(* IEC 61131-3 sources: Lasal-MCP/examples/SampleSource/LASALScreenAdvancedSolution/LASALScreenAdvancedSolution/LASALScreenAdvacnedSolution/Stations/Terminal/HMI/Class/InputMyIO, 1 file *)

(* ---- InputMyIO.st ---- *)
#define CROSSHAIR_LENGTH 20
#define CROSSHAIR_WIDTH 1
#define OFFSET_X 10
#define OFFSET_Y 5

(*!
<Class
	Name               = "InputMyIO"
	Revision           = "0.0"
	RealtimeTask       = "false"
	CyclicTask         = "false"
	BackgroundTask     = "false"
	Sigmatek           = "false"
	OSInterface        = "false"
	HighPriority       = "false"
	Automatic          = "false"
	UpdateMode         = "Prescan"
	SharedCommandTable = "true"
	Objectsize         = "(450,300)">
	<Channels>
		<Server Name="CoordX" Visualized="true" Initialize="false" WriteProtected="false" Retentive="false"/>
		<Server Name="CoordY" Visualized="true" Initialize="false" WriteProtected="false" Retentive="false"/>
		<Client Name="_Grafix" Required="false" Internal="false"/>
	</Channels>
	<Network Name="InputMyIO">
		<!-- List of Components in this network -->
		<Components>
			<Object
				Name       = "_base"
				Class      = "_MyIO"
				Position   = "(218,120)"
				Visualized = "true"
				Remotely   = "true">
				<Channels>
					<Server Name="Refresh"/>
					<Server Name="Server0"/>
					<Client Name="Graphic"/>
					<Client Name="Lse"/>
				</Channels>
			</Object>
		</Components>
		<Comments>
		</Comments>
		<!-- List of Connections in this network -->
		<Connections>
			<Connection Source="this.Server0" Destination="_base.Server0" Vertices="(706,210),(534,210),"/>
			<Connection Source="this.Refresh" Destination="_base.Refresh" Vertices="(706,270),(534,270),"/>
			<Connection Source="_base.Lse" Destination="this.Lse" Vertices="(218,210),(38,210),"/>
		</Connections>
		<!-- Headerfiles -->
		<Options>
		</Options>
	</Network>
</Class>
*)
#pragma using _MyIO

InputMyIO : CLASS
: _MyIO
  //Servers:
	CoordX 	: SvrCh_DINT;
	CoordY 	: SvrCh_DINT;
  //Clients:
	_Grafix 	: CltChCmd__Grafix;
  //Variables:
		myFocus 	: BOOL;
  //Functions:
				//! <Function Comment="this method will be called once when the focus will be given to this object" Name="GetFocus"/>
	FUNCTION __CDECL VIRTUAL GLOBAL GetFocus
		VAR_INPUT
			pio 	: ^_IO;			//! <Variable Comment="pointer to _IO information" Name="GetFocus.pio"/>
		END_VAR
		VAR_OUTPUT
			retcode (EAX) 	: _DOIT;			//! <Variable Comment="return _IFAILED if you dont want to get the focus on the other hand _IDLE" Name="GetFocus.retcode"/>
		END_VAR;
				//! <Function Comment="this method is called once when the focus is taken from object" Name="KillFocus"/>
	FUNCTION __CDECL VIRTUAL GLOBAL KillFocus
		VAR_INPUT
			pio 	: ^_IO;			//! <Variable Comment="pointer to _IO information" Name="KillFocus.pio"/>
		END_VAR
		VAR_OUTPUT
			retcode (EAX) 	: _DOIT;			//! <Variable Comment="return always _IDLE because you can&apos;t prevent action" Name="KillFocus.retcode"/>
		END_VAR;
				//! <Function Comment="this method is called everytime when the input is active and a event occured" Name="GetEvent"/>
	FUNCTION __CDECL VIRTUAL GLOBAL GetEvent
		VAR_INPUT
			ped 	: ^_EDITOR;			//! <Variable Comment="pointer to _EDITOR information" Name="GetEvent.ped"/>
			pe 	: ^_EVENT;			//! <Variable Comment="pointer to _EVENT information" Name="GetEvent.pe"/>
		END_VAR
		VAR_OUTPUT
			retcode (EAX) 	: _DOIT;			//! <Variable Comment="for the returnstatement there are 3 different possibilities&#13;&#10;  _IDLE ..... the system should goon like it is (system goes on)&#13;&#10;  _IDIDIT ... i did it (system is ready)&#13;&#10;  _IFAILED .. i tried to do my best, but i failed (system is ready)&#13;&#10;" Name="GetEvent.retcode"/>
		END_VAR;
				//! <Function Comment="this method is called everytime when system wants to redraw the io" Name="Draw"/>
	FUNCTION __CDECL VIRTUAL GLOBAL Draw
		VAR_INPUT
			pio 	: ^_IO;			//! <Variable Comment="pointer to _IO information" Name="Draw.pio"/>
			pr 	: ^_RESULT;			//! <Variable Comment="pointer to _RESULT information" Name="Draw.pr"/>
			pv 	: ^_VARIABLE;			//! <Variable Comment="pointer to io _VARIABLE information" Name="Draw.pv"/>
			input 	: BOOL;			//! <Variable Comment="TRUE it&apos;s an input&#13;&#10;FALSE it&apos;s an output" Name="Draw.input"/>
		END_VAR
		VAR_OUTPUT
			retcode (EAX) 	: _DOIT;			//! <Variable Comment="for the returnstatement there are 3 different possibilities&#13;&#10;  _IDLE ..... the system should goon like it is (system goes on)&#13;&#10;  _IDIDIT ... i did it (system is ready)&#13;&#10;  _IFAILED .. i tried to do my best, but i failed (system is re" Name="Draw.retcode"/>
		END_VAR;
				//! <Function Comment="this method is called everytime when system wants to get data for defined io.&#13;&#10;&#13;&#10;pr ........ &#13;&#10;pio ....... pointer to io information&#13;&#10;pv ........ pointer to io variableinformation&#13;&#10;input ..... TRUE it&apos;s an input / FALSE it&apos;s an output&#13;&#10;&#13;&#10;for the returnstatement there are 3 different possibilities&#13;&#10;_IDLE ..... the system should goon like it is (system goes on)&#13;&#10;_IDIDIT ... i did it (system is ready)&#13;&#10;_IFAILED .. i tried to do my best, but i failed (system is ready)&#13;&#10;&#13;&#10;if you want to do it let&apos;s return _IDIDIT and initialize the  structure _RESULT&#13;&#10;" Name="GetData"/>
	FUNCTION __CDECL VIRTUAL GLOBAL GetData
		VAR_INPUT
			pr 	: ^_RESULT;			//! <Variable Comment="pointer to _RESULT information" Name="GetData.pr"/>
			pio 	: ^_IO;			//! <Variable Comment="pointer to _IO information" Name="GetData.pio"/>
			pv 	: ^_VARIABLE;			//! <Variable Comment="pointer to _VARIABLE information given by LSE" Name="GetData.pv"/>
			input 	: BOOL;			//! <Variable Comment="TRUE it&apos;s an input&#13;&#10;FALSE it&apos;s an output" Name="GetData.input"/>
		END_VAR
		VAR_OUTPUT
			retcode (EAX) 	: _DOIT;			//! <Variable Comment="for the returnstatement there are 3 different possibilities&#13;&#10;  _IDLE ..... the system should goon like it is (system goes on)&#13;&#10;  _IDIDIT ... i did it (system is ready)&#13;&#10;  _IFAILED .. i tried to do my best, but i failed (system is ready)" Name="GetData.retcode"/>
		END_VAR;
				//! <Function Comment="this method is called once right in front of drawing the object.&#13;&#10;for example open screen&#13;&#10;" Name="IF_Start"/>
	FUNCTION __CDECL VIRTUAL GLOBAL IF_Start
		VAR_INPUT
			pio 	: ^_IO;			//! <Variable Comment="pointer to _IO information" Name="IF_Start.pio"/>
			firsttime 	: BOOL;			//! <Variable Comment="true: when system wants to view drawing after open screen&#13;&#10;false: when system wants to redraw background" Name="IF_Start.firsttime"/>
		END_VAR;
  //Tables:
	FUNCTION @STD
		VAR_OUTPUT
			ret_code	: CONFSTATES;
		END_VAR;
	FUNCTION GLOBAL TAB @CT_;
END_CLASS;

#pragma usingLtd _Grafix

FUNCTION __CDECL VIRTUAL GLOBAL InputMyIO::IF_Start
	VAR_INPUT
		pio 	: ^_IO;
		firsttime 	: BOOL;
	END_VAR

  _MyIO::IF_Start(pio:= pio, firsttime:= firsttime);

  if (firsttime = TRUE) then

    CoordX := (pio^.room.xy2.x - pio^.room.xy1.x) / 2;
    CoordY := (pio^.room.xy2.y - pio^.room.xy1.y) / 2;

  end_if;

END_FUNCTION

FUNCTION __CDECL VIRTUAL GLOBAL InputMyIO::GetData
	VAR_INPUT
		pr 	: ^_RESULT;
		pio 	: ^_IO;
		pv 	: ^_VARIABLE;
		input 	: BOOL;
	END_VAR
	VAR_OUTPUT
		retcode (EAX) 	: _DOIT;
	END_VAR

  _MyIO::GetData(pr:= pr, pio:= pio, pv:= pv, input:= input);

  pr^.value := to_dint((to_udint(CoordX) rol 1) xor (to_udint(CoordY)));

  retcode := _IDIDIT;

END_FUNCTION

FUNCTION __CDECL VIRTUAL GLOBAL InputMyIO::GetEvent
	VAR_INPUT
		ped 	: ^_EDITOR;
		pe 	: ^_EVENT;
	END_VAR
	VAR_OUTPUT
		retcode (EAX) 	: _DOIT;
	END_VAR

  retcode := _IDLE;

  if ((pe^.ftype = _EVENT_HIDMOVE) | (pe^.ftype = _EVENT_HIDPRESS)) then

    if ((pe^.dot.x >= ped^.input.io.space.xy1.x) &
        (pe^.dot.x <= ped^.input.io.space.xy2.x) &
        (pe^.dot.y >= ped^.input.io.space.xy1.y) &
        (pe^.dot.y <= ped^.input.io.space.xy2.y))
    then

      CoordX := pe^.dot.x - ped^.input.io.space.xy1.x;
      CoordY := pe^.dot.y - ped^.input.io.space.xy1.y;

      retcode := _IDIDIT;

    end_if;

  end_if;

END_FUNCTION

FUNCTION __CDECL VIRTUAL GLOBAL InputMyIO::GetFocus
	VAR_INPUT
		pio 	: ^_IO;
	END_VAR
	VAR_OUTPUT
		retcode (EAX) 	: _DOIT;
	END_VAR

  _MyIO::GetFocus(pio:=pio);

  myFocus := TRUE;
  retcode := _IDIDIT;

END_FUNCTION

FUNCTION __CDECL VIRTUAL GLOBAL InputMyIO::KillFocus
	VAR_INPUT
		pio 	: ^_IO;
	END_VAR
	VAR_OUTPUT
		retcode (EAX) 	: _DOIT;
	END_VAR

  _MyIO::KillFocus(pio:=pio);

  myFocus := FALSE;
  retcode := _IDIDIT;

END_FUNCTION

FUNCTION __CDECL VIRTUAL GLOBAL InputMyIO::Draw
	VAR_INPUT
		pio 	: ^_IO;
		pr 	: ^_RESULT;
		pv 	: ^_VARIABLE;
		input 	: BOOL;
	END_VAR
	VAR_OUTPUT
		retcode (EAX) 	: _DOIT;
	END_VAR
  VAR
    act : _NEWSCREEN;
    x : _KOORD;
    y : _KOORD;
    color : _COLOR;
    xText : array[0..6] of char;
    yText : array[0..6] of char;
    xAttribute : _ATTRIB;
    yAttribute : _ATTRIB;
    xTextPos : _DOT;
    yTextPos : _DOT;
  END_VAR

  push_screen(p0:= #act);

  _Grafix.PutImage(image:= #pio^.image, x0:= DEFKOORD, y0:= DEFKOORD);

  x := to_int(CoordX) + pio^.space.xy1.x;
  y := to_int(CoordY) + pio^.space.xy1.y;

  if (myFocus = TRUE) then
    color := GetEditColorBack(x0:= _EDITACTIVE);
  else
    color := pio^.coltxt;
  end_if;

  // set alignment and position for koord values to display
  if (CoordX < (pio^.space.xy2.x - pio^.space.xy1.x) / 2) then
    xAttribute := T_LEFTBOUND;
    yAttribute := T_RIGHTBOUND;
    xTextPos.x := x + OFFSET_X;
    yTextPos.x := pio^.space.xy2.x - OFFSET_X;
  else
    xAttribute := T_RIGHTBOUND;
    yAttribute := T_LEFTBOUND;
    xTextPos.x := x - OFFSET_X;
    yTextPos.x := pio^.space.xy1.x + OFFSET_X;
  end_if;

  if (CoordY < (pio^.space.xy2.y - pio^.space.xy1.y) / 2) then
    xAttribute := xAttribute or T_DOWNBOUND;
    xTextPos.y := pio^.space.xy2.y - OFFSET_Y;
    yTextPos.y := y + OFFSET_Y;
  else
    yAttribute := yAttribute or T_DOWNBOUND;
    xTextPos.y := pio^.space.xy1.y + OFFSET_Y;
    yTextPos.y := y - OFFSET_Y;
  end_if;

  // draw frame
  _Grafix.Rectangle(x0:= pio^.space.xy1.x,
                    y0:= pio^.space.xy1.y,
                    x1:= pio^.space.xy2.x,
                    y1:= pio^.space.xy2.y,
                    attrib:= pio^.attrib,
                    color:= pio^.colframe);

  // draw horizontal line
  _Grafix.Line(x0:= pio^.space.xy1.x + 1,
               y0:= y,
               x1:= pio^.space.xy2.x - 1,
               y1:= y,
               attrib:= pio^.attrib,
               color:= color);

  // draw vertical line
  _Grafix.Line(x0:= x,
               y0:= pio^.space.xy1.y + 1,
               x1:= x,
               y1:= pio^.space.xy2.y - 1,
               attrib:= pio^.attrib,
               color:= color);

  // draw crosshair in the middle
  _Grafix.Beam(x0:= x - CROSSHAIR_LENGTH,
               y0:= y - CROSSHAIR_WIDTH,
               x1:= x + CROSSHAIR_LENGTH,
               y1:= y + CROSSHAIR_WIDTH,
               attrib:= pio^.attrib,
               color:= color);

  _Grafix.Beam(x0:= x - CROSSHAIR_WIDTH,
               y0:= y - CROSSHAIR_LENGTH,
               x1:= x + CROSSHAIR_WIDTH,
               y1:= y + CROSSHAIR_LENGTH,
               attrib:= pio^.attrib,
               color:= color);

  // convert value into string
  DToA(p0:= #xText[0],
       x1:= CoordX,
       x2:= 16#0800,
       x3:= sizeof(_ASCII));

  DToA(p0:= #yText[0],
       x1:= CoordY,
       x2:= 16#0800,
       x3:= sizeof(_ASCII));

  // draw koords on right position
  _Grafix.OutTextXY(x0:= xTextPos.x,
                    y0:= xTextPos.y,
                    textptr:= #xText[0],
                    attrib:= xAttribute,
                    color:= _Grafix.MakeColor(backcolor:= INVISIBLE, frontcolor:= WHITE),
                    chr_size:=sizeof(_ASCII));

  _Grafix.OutTextXY(x0:= yTextPos.x,
                    y0:= yTextPos.y,
                    textptr:= #yText[0],
                    attrib:= yAttribute,
                    color:= _Grafix.MakeColor(backcolor:= INVISIBLE, frontcolor:= WHITE),
                    chr_size:= sizeof(_ASCII));

  pop_screen(p0:= #act);
  copy_screen(p0:= #act, p1:= #pio^.space);

  retcode := _IDIDIT;

END_FUNCTION
